// TIA Portal project "039_fw41" (V21)

(* hardware
DEVICE "PLC_1"  S7-1500 station
   slot 0: "Rail_0"  Rack  6ES7 590-1***0-0AA0
   slot 1: "PLC_1"  CPU 1516-3 PN/DP  6ES7 516-3AP03-0AB0  V4.1
      slot 3: "CPU display_1"  6ES7591-1BA00-0AA0
      slot 32768: "PROFINET interface_1"  X1
         slot 32769: "Port_1"  X1 P1
         slot 32770: "Port_2"  X1 P2
      slot 33024: "PROFINET interface_2"  X2
         slot 33025: "Port_1"  X2 P1
      slot 33280: "DP interface_1"  X3
      slot 34817: "Virtual CP interface port_1"  Virtual CP interface port  Virtual CP interface port FW V4.1
*)

// ===== PLC "PLC_1"  CPU 1516-3 PN/DP =====

DATA_BLOCK "DB_Arr"   // DB1
{ S7_Optimized_Access := 'FALSE' }
   VAR
      "a" : Array[0..9] of Int;
      "b" : Array[0..9] of Int;
      w : Array[0..3] of Word;
      r : Array[0..3] of Real;
      "by" : Array[0..7] of Byte;
      bits : Array[0..15] of Bool;
   END_VAR
BEGIN
END_DATA_BLOCK

FUNCTION_BLOCK "FX_Lad_103"   // FB1, LAD
{ S7_Optimized_Access := 'TRUE' }
VERSION : 0.1
   VAR_INPUT
      "a" : Bool;
      "b" : Bool;
      c : Bool;
      ia : Int;
      ib : Int;
      ic : Int;
      da : DInt;
      db : DInt;
      ra : Real;
      rb : Real;
      wa : Word;
      wb : Word;
      dwa : DWord;
      ba : Byte;
      ta : Time;
      tb : Time;
      s1 : String;
      s2 : String;
   END_VAR
   VAR_OUTPUT
      q : Bool;
      q2 : Bool;
      io : Int;
      io2 : Int;
      dout : DInt;
      rout : Real;
      wout : Word;
      dwout : DWord;
      bout : Byte;
      tout : Time;
      sout : String;
   END_VAR
   VAR_IN_OUT
      x_bool : Bool;
      x_uint : UInt;
      arr : Array[0..9] of Int;
      barr : Array[0..7] of Bool;
      iinout : Int;
   END_VAR
   VAR
      ton1 : TON_TIME;
      tof1 : TOF_TIME;
      tp1 : TP_TIME;
      tonr1 : TONR_TIME;
      ctu1 : CTU_INT;
      ctd1 : CTD_INT;
      ctud1 : CTUD_INT;
      rtrig1 : R_TRIG;
      ftrig1 : F_TRIG;
      edge1 : Bool;
      edge2 : Bool;
      stat1 : Bool;
      stat2 : Bool;
      stati : Int;
   END_VAR
   VAR_TEMP
      t1 : Bool;
      t2 : Bool;
      ti : Int;
      td : DInt;
      tr : Real;
      tw : Word;
      tt : Time;
      var1 : Variant;
   END_VAR
BEGIN

REGION Network 1: ---| |--- - Normally open contact
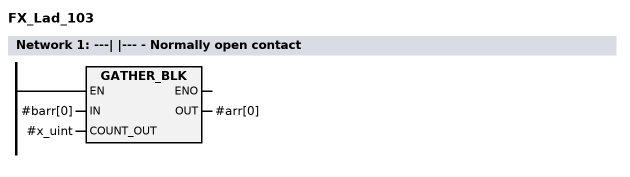
   GATHER_BLK(IN := #barr[0], COUNT_OUT := #x_uint, OUT => #arr[0]);
END_REGION
END_FUNCTION_BLOCK

FUNCTION_BLOCK "FX_TP2"   // FB2, LAD
{ S7_Optimized_Access := 'TRUE' }
VERSION : 0.1
   VAR_INPUT
      "a" : Bool;
      "b" : Bool;
      c : Bool;
      ia : Int;
      ib : Int;
      ic : Int;
      da : DInt;
      db : DInt;
      ra : Real;
      rb : Real;
      wa : Word;
      wb : Word;
      dwa : DWord;
      ba : Byte;
      ta : Time;
      tb : Time;
      s1 : String;
      s2 : String;
   END_VAR
   VAR_OUTPUT
      q : Bool;
      q2 : Bool;
      io : Int;
      io2 : Int;
      dout : DInt;
      rout : Real;
      wout : Word;
      dwout : DWord;
      bout : Byte;
      tout : Time;
      sout : String;
   END_VAR
   VAR_IN_OUT
      arr : Array[0..9] of Int;
      barr : Array[0..7] of Bool;
      iinout : Int;
   END_VAR
   VAR
      ton1 : TON_TIME;
      tof1 : TOF_TIME;
      tp1 : TP_TIME;
      tonr1 : TONR_TIME;
      ctu1 : CTU_INT;
      ctd1 : CTD_INT;
      ctud1 : CTUD_INT;
      rtrig1 : R_TRIG;
      ftrig1 : F_TRIG;
      edge1 : Bool;
      edge2 : Bool;
      stat1 : Bool;
      stat2 : Bool;
      stati : Int;
   END_VAR
   VAR_TEMP
      t1 : Bool;
      t2 : Bool;
      ti : Int;
      td : DInt;
      tr : Real;
      tw : Word;
      tt : Time;
      var1 : Variant;
   END_VAR
BEGIN

REGION Network 1: ---| |--- - Normally open contact
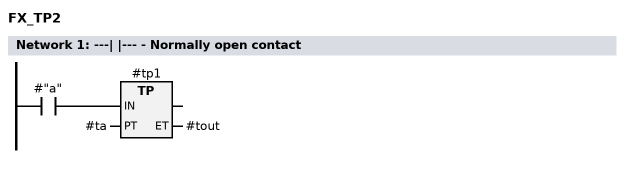
   #tp1(IN := #"a", PT := #ta, ET => #tout);   // TP
END_REGION
END_FUNCTION_BLOCK

FUNCTION_BLOCK "FX_Lad_024"   // FB3, LAD
{ S7_Optimized_Access := 'TRUE' }
VERSION : 0.1
   VAR_INPUT
      "a" : Bool;
      "b" : Bool;
      c : Bool;
      ia : Int;
      ib : Int;
      ic : Int;
      da : DInt;
      db : DInt;
      ra : Real;
      rb : Real;
      wa : Word;
      wb : Word;
      dwa : DWord;
      ba : Byte;
      ta : Time;
      tb : Time;
      s1 : String;
      s2 : String;
   END_VAR
   VAR_OUTPUT
      q : Bool;
      q2 : Bool;
      io : Int;
      io2 : Int;
      dout : DInt;
      rout : Real;
      wout : Word;
      dwout : DWord;
      bout : Byte;
      tout : Time;
      sout : String;
   END_VAR
   VAR_IN_OUT
      arr : Array[0..9] of Int;
      barr : Array[0..7] of Bool;
      iinout : Int;
   END_VAR
   VAR
      ton1 : TON_TIME;
      tof1 : TOF_TIME;
      tp1 : TP_TIME;
      tonr1 : TONR_TIME;
      ctu1 : CTU_INT;
      ctd1 : CTD_INT;
      ctud1 : CTUD_INT;
      rtrig1 : R_TRIG;
      ftrig1 : F_TRIG;
      edge1 : Bool;
      edge2 : Bool;
      stat1 : Bool;
      stat2 : Bool;
      stati : Int;
   END_VAR
   VAR_TEMP
      t1 : Bool;
      t2 : Bool;
      ti : Int;
      td : DInt;
      tr : Real;
      tw : Word;
      tt : Time;
      var1 : Variant;
   END_VAR
BEGIN

REGION Network 1: ---| |--- - Normally open contact
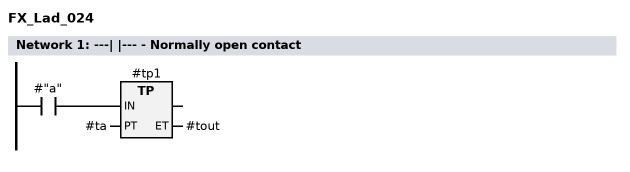
   #tp1(IN := #"a", PT := #ta, ET => #tout);   // TP
END_REGION
END_FUNCTION_BLOCK

FUNCTION_BLOCK "FX_Lad_025"   // FB4, LAD
{ S7_Optimized_Access := 'TRUE' }
VERSION : 0.1
   VAR_INPUT
      "a" : Bool;
      "b" : Bool;
      c : Bool;
      ia : Int;
      ib : Int;
      ic : Int;
      da : DInt;
      db : DInt;
      ra : Real;
      rb : Real;
      wa : Word;
      wb : Word;
      dwa : DWord;
      ba : Byte;
      ta : Time;
      tb : Time;
      s1 : String;
      s2 : String;
   END_VAR
   VAR_OUTPUT
      q : Bool;
      q2 : Bool;
      io : Int;
      io2 : Int;
      dout : DInt;
      rout : Real;
      wout : Word;
      dwout : DWord;
      bout : Byte;
      tout : Time;
      sout : String;
   END_VAR
   VAR_IN_OUT
      arr : Array[0..9] of Int;
      barr : Array[0..7] of Bool;
      iinout : Int;
   END_VAR
   VAR
      ton1 : TON_TIME;
      tof1 : TOF_TIME;
      tp1 : TP_TIME;
      tonr1 : TONR_TIME;
      ctu1 : CTU_INT;
      ctd1 : CTD_INT;
      ctud1 : CTUD_INT;
      rtrig1 : R_TRIG;
      ftrig1 : F_TRIG;
      edge1 : Bool;
      edge2 : Bool;
      stat1 : Bool;
      stat2 : Bool;
      stati : Int;
   END_VAR
   VAR_TEMP
      t1 : Bool;
      t2 : Bool;
      ti : Int;
      td : DInt;
      tr : Real;
      tw : Word;
      tt : Time;
      var1 : Variant;
   END_VAR
BEGIN

REGION Network 1: ---| |--- - Normally open contact
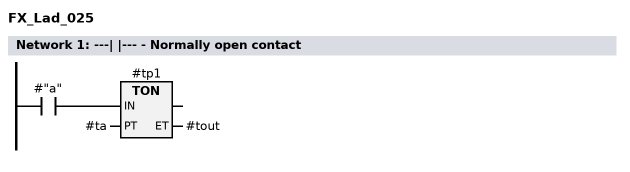
   #tp1(IN := #"a", PT := #ta, ET => #tout);   // TON
END_REGION
END_FUNCTION_BLOCK

FUNCTION_BLOCK "FX_Lad_026"   // FB5, LAD
{ S7_Optimized_Access := 'TRUE' }
VERSION : 0.1
   VAR_INPUT
      "a" : Bool;
      "b" : Bool;
      c : Bool;
      ia : Int;
      ib : Int;
      ic : Int;
      da : DInt;
      db : DInt;
      ra : Real;
      rb : Real;
      wa : Word;
      wb : Word;
      dwa : DWord;
      ba : Byte;
      ta : Time;
      tb : Time;
      s1 : String;
      s2 : String;
   END_VAR
   VAR_OUTPUT
      q : Bool;
      q2 : Bool;
      io : Int;
      io2 : Int;
      dout : DInt;
      rout : Real;
      wout : Word;
      dwout : DWord;
      bout : Byte;
      tout : Time;
      sout : String;
   END_VAR
   VAR_IN_OUT
      arr : Array[0..9] of Int;
      barr : Array[0..7] of Bool;
      iinout : Int;
   END_VAR
   VAR
      ton1 : TON_TIME;
      tof1 : TOF_TIME;
      tp1 : TP_TIME;
      tonr1 : TONR_TIME;
      ctu1 : CTU_INT;
      ctd1 : CTD_INT;
      ctud1 : CTUD_INT;
      rtrig1 : R_TRIG;
      ftrig1 : F_TRIG;
      edge1 : Bool;
      edge2 : Bool;
      stat1 : Bool;
      stat2 : Bool;
      stati : Int;
   END_VAR
   VAR_TEMP
      t1 : Bool;
      t2 : Bool;
      ti : Int;
      td : DInt;
      tr : Real;
      tw : Word;
      tt : Time;
      var1 : Variant;
   END_VAR
BEGIN

REGION Network 1: ---| |--- - Normally open contact
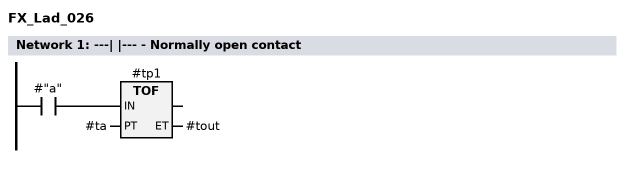
   #tp1(IN := #"a", PT := #ta, ET => #tout);   // TOF
END_REGION
END_FUNCTION_BLOCK

FUNCTION_BLOCK "FX_Lad_027"   // FB6, LAD
{ S7_Optimized_Access := 'TRUE' }
VERSION : 0.1
   VAR_INPUT
      "a" : Bool;
      "b" : Bool;
      c : Bool;
      ia : Int;
      ib : Int;
      ic : Int;
      da : DInt;
      db : DInt;
      ra : Real;
      rb : Real;
      wa : Word;
      wb : Word;
      dwa : DWord;
      ba : Byte;
      ta : Time;
      tb : Time;
      s1 : String;
      s2 : String;
   END_VAR
   VAR_OUTPUT
      q : Bool;
      q2 : Bool;
      io : Int;
      io2 : Int;
      dout : DInt;
      rout : Real;
      wout : Word;
      dwout : DWord;
      bout : Byte;
      tout : Time;
      sout : String;
   END_VAR
   VAR_IN_OUT
      arr : Array[0..9] of Int;
      barr : Array[0..7] of Bool;
      iinout : Int;
   END_VAR
   VAR
      ton1 : TON_TIME;
      tof1 : TOF_TIME;
      tp1 : TP_TIME;
      tonr1 : TONR_TIME;
      ctu1 : CTU_INT;
      ctd1 : CTD_INT;
      ctud1 : CTUD_INT;
      rtrig1 : R_TRIG;
      ftrig1 : F_TRIG;
      edge1 : Bool;
      edge2 : Bool;
      stat1 : Bool;
      stat2 : Bool;
      stati : Int;
   END_VAR
   VAR_TEMP
      t1 : Bool;
      t2 : Bool;
      ti : Int;
      td : DInt;
      tr : Real;
      tw : Word;
      tt : Time;
      var1 : Variant;
   END_VAR
BEGIN

REGION Network 1: ---| |--- - Normally open contact
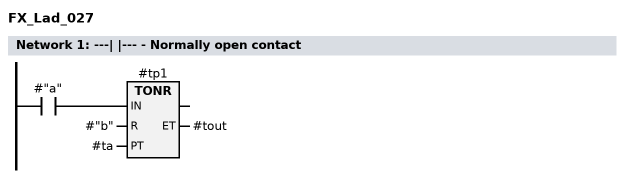
   #tp1(IN := #"a", R := #"b", PT := #ta, ET => #tout);   // TONR
END_REGION
END_FUNCTION_BLOCK

FUNCTION_BLOCK "FX_Lad_ex003"   // FB7, LAD
{ S7_Optimized_Access := 'TRUE' }
VERSION : 0.1
   VAR_INPUT
      "a" : Bool;
      "b" : Bool;
      c : Bool;
      ia : Int;
      ib : Int;
      ic : Int;
      da : DInt;
      db : DInt;
      ra : Real;
      rb : Real;
      wa : Word;
      wb : Word;
      dwa : DWord;
      ba : Byte;
      ta : Time;
      tb : Time;
      s1 : String;
      s2 : String;
   END_VAR
   VAR_OUTPUT
      q : Bool;
      q2 : Bool;
      io : Int;
      io2 : Int;
      dout : DInt;
      rout : Real;
      wout : Word;
      dwout : DWord;
      bout : Byte;
      tout : Time;
      sout : String;
   END_VAR
   VAR_IN_OUT
      x_time : Time;
      arr : Array[0..9] of Int;
      barr : Array[0..7] of Bool;
      iinout : Int;
   END_VAR
   VAR
      ton1 : TON_TIME;
      tof1 : TOF_TIME;
      tp1 : TP_TIME;
      tonr1 : TONR_TIME;
      ctu1 : CTU_INT;
      ctd1 : CTD_INT;
      ctud1 : CTUD_INT;
      rtrig1 : R_TRIG;
      ftrig1 : F_TRIG;
      edge1 : Bool;
      edge2 : Bool;
      stat1 : Bool;
      stat2 : Bool;
      stati : Int;
   END_VAR
   VAR_TEMP
      t1 : Bool;
      t2 : Bool;
      ti : Int;
      td : DInt;
      tr : Real;
      tw : Word;
      tt : Time;
      var1 : Variant;
   END_VAR
BEGIN

REGION Network 1: ---| |--- - Normally open contact
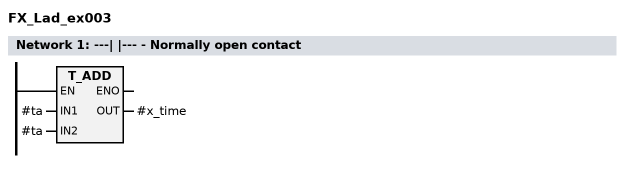
   #x_time := T_ADD(IN1 := #ta, IN2 := #ta);
END_REGION
END_FUNCTION_BLOCK

FUNCTION_BLOCK "FX_Lad_ex004"   // FB8, LAD
{ S7_Optimized_Access := 'TRUE' }
VERSION : 0.1
   VAR_INPUT
      "a" : Bool;
      "b" : Bool;
      c : Bool;
      ia : Int;
      ib : Int;
      ic : Int;
      da : DInt;
      db : DInt;
      ra : Real;
      rb : Real;
      wa : Word;
      wb : Word;
      dwa : DWord;
      ba : Byte;
      ta : Time;
      tb : Time;
      s1 : String;
      s2 : String;
   END_VAR
   VAR_OUTPUT
      q : Bool;
      q2 : Bool;
      io : Int;
      io2 : Int;
      dout : DInt;
      rout : Real;
      wout : Word;
      dwout : DWord;
      bout : Byte;
      tout : Time;
      sout : String;
   END_VAR
   VAR_IN_OUT
      x_time : Time;
      arr : Array[0..9] of Int;
      barr : Array[0..7] of Bool;
      iinout : Int;
   END_VAR
   VAR
      ton1 : TON_TIME;
      tof1 : TOF_TIME;
      tp1 : TP_TIME;
      tonr1 : TONR_TIME;
      ctu1 : CTU_INT;
      ctd1 : CTD_INT;
      ctud1 : CTUD_INT;
      rtrig1 : R_TRIG;
      ftrig1 : F_TRIG;
      edge1 : Bool;
      edge2 : Bool;
      stat1 : Bool;
      stat2 : Bool;
      stati : Int;
   END_VAR
   VAR_TEMP
      t1 : Bool;
      t2 : Bool;
      ti : Int;
      td : DInt;
      tr : Real;
      tw : Word;
      tt : Time;
      var1 : Variant;
   END_VAR
BEGIN

REGION Network 1: ---| |--- - Normally open contact
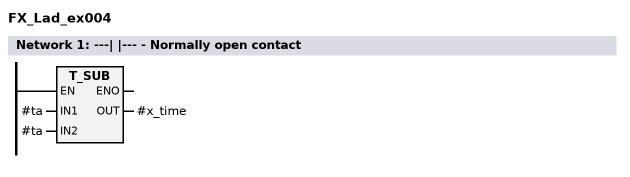
   #x_time := T_SUB(IN1 := #ta, IN2 := #ta);
END_REGION
END_FUNCTION_BLOCK

FUNCTION_BLOCK "FX_Lad_ex018"   // FB9, LAD
{ S7_Optimized_Access := 'TRUE' }
VERSION : 0.1
   VAR_INPUT
      "a" : Bool;
      "b" : Bool;
      c : Bool;
      ia : Int;
      ib : Int;
      ic : Int;
      da : DInt;
      db : DInt;
      ra : Real;
      rb : Real;
      wa : Word;
      wb : Word;
      dwa : DWord;
      ba : Byte;
      ta : Time;
      tb : Time;
      s1 : String;
      s2 : String;
   END_VAR
   VAR_OUTPUT
      q : Bool;
      q2 : Bool;
      io : Int;
      io2 : Int;
      dout : DInt;
      rout : Real;
      wout : Word;
      dwout : DWord;
      bout : Byte;
      tout : Time;
      sout : String;
   END_VAR
   VAR_IN_OUT
      arr : Array[0..9] of Int;
      barr : Array[0..7] of Bool;
      iinout : Int;
   END_VAR
   VAR
      ton1 : TON_TIME;
      tof1 : TOF_TIME;
      tp1 : TP_TIME;
      tonr1 : TONR_TIME;
      ctu1 : CTU_INT;
      ctd1 : CTD_INT;
      ctud1 : CTUD_INT;
      rtrig1 : R_TRIG;
      ftrig1 : F_TRIG;
      edge1 : Bool;
      edge2 : Bool;
      stat1 : Bool;
      stat2 : Bool;
      stati : Int;
   END_VAR
   VAR_TEMP
      t1 : Bool;
      t2 : Bool;
      ti : Int;
      td : DInt;
      tr : Real;
      tw : Word;
      tt : Time;
      var1 : Variant;
   END_VAR
BEGIN

REGION Network 1: ---| |--- - Normally open contact
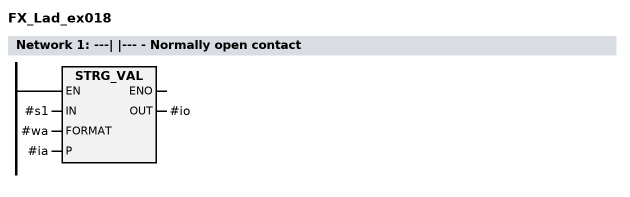
   STRG_VAL(IN := #s1, FORMAT := #wa, P := #ia, OUT => #io);
END_REGION
END_FUNCTION_BLOCK

FUNCTION_BLOCK "FX_Lad_ex019"   // FB10, LAD
{ S7_Optimized_Access := 'TRUE' }
VERSION : 0.1
   VAR_INPUT
      "a" : Bool;
      "b" : Bool;
      c : Bool;
      ia : Int;
      ib : Int;
      ic : Int;
      da : DInt;
      db : DInt;
      ra : Real;
      rb : Real;
      wa : Word;
      wb : Word;
      dwa : DWord;
      ba : Byte;
      ta : Time;
      tb : Time;
      s1 : String;
      s2 : String;
   END_VAR
   VAR_OUTPUT
      q : Bool;
      q2 : Bool;
      io : Int;
      io2 : Int;
      dout : DInt;
      rout : Real;
      wout : Word;
      dwout : DWord;
      bout : Byte;
      tout : Time;
      sout : String;
   END_VAR
   VAR_IN_OUT
      arr : Array[0..9] of Int;
      barr : Array[0..7] of Bool;
      iinout : Int;
   END_VAR
   VAR
      ton1 : TON_TIME;
      tof1 : TOF_TIME;
      tp1 : TP_TIME;
      tonr1 : TONR_TIME;
      ctu1 : CTU_INT;
      ctd1 : CTD_INT;
      ctud1 : CTUD_INT;
      rtrig1 : R_TRIG;
      ftrig1 : F_TRIG;
      edge1 : Bool;
      edge2 : Bool;
      stat1 : Bool;
      stat2 : Bool;
      stati : Int;
   END_VAR
   VAR_TEMP
      t1 : Bool;
      t2 : Bool;
      ti : Int;
      td : DInt;
      tr : Real;
      tw : Word;
      tt : Time;
      var1 : Variant;
   END_VAR
BEGIN

REGION Network 1: ---| |--- - Normally open contact
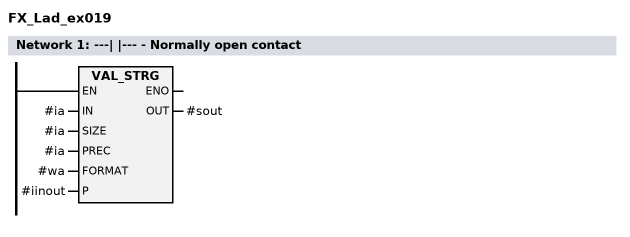
   VAL_STRG(IN := #ia, SIZE := #ia, PREC := #ia, FORMAT := #wa, P := #iinout, OUT => #sout);
END_REGION
END_FUNCTION_BLOCK

FUNCTION_BLOCK "FX_Lad_ex021"   // FB11, LAD
{ S7_Optimized_Access := 'TRUE' }
VERSION : 0.1
   VAR_INPUT
      "a" : Bool;
      "b" : Bool;
      c : Bool;
      ia : Int;
      ib : Int;
      ic : Int;
      da : DInt;
      db : DInt;
      ra : Real;
      rb : Real;
      wa : Word;
      wb : Word;
      dwa : DWord;
      ba : Byte;
      ta : Time;
      tb : Time;
      s1 : String;
      s2 : String;
   END_VAR
   VAR_OUTPUT
      q : Bool;
      q2 : Bool;
      io : Int;
      io2 : Int;
      dout : DInt;
      rout : Real;
      wout : Word;
      dwout : DWord;
      bout : Byte;
      tout : Time;
      sout : String;
   END_VAR
   VAR_IN_OUT
      x_variant : Variant;
      arr : Array[0..9] of Int;
      barr : Array[0..7] of Bool;
      iinout : Int;
   END_VAR
   VAR
      ton1 : TON_TIME;
      tof1 : TOF_TIME;
      tp1 : TP_TIME;
      tonr1 : TONR_TIME;
      ctu1 : CTU_INT;
      ctd1 : CTD_INT;
      ctud1 : CTUD_INT;
      rtrig1 : R_TRIG;
      ftrig1 : F_TRIG;
      edge1 : Bool;
      edge2 : Bool;
      stat1 : Bool;
      stat2 : Bool;
      stati : Int;
   END_VAR
   VAR_TEMP
      t1 : Bool;
      t2 : Bool;
      ti : Int;
      td : DInt;
      tr : Real;
      tw : Word;
      tt : Time;
      var1 : Variant;
   END_VAR
BEGIN

REGION Network 1: ---| |--- - Normally open contact
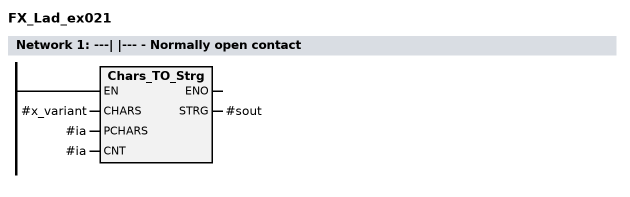
   // no SCL statement known for Chars_TO_Strg: written as a call
   Chars_TO_Strg(Chars := #x_variant, pChars := #ia, Cnt := #ia, Strg => #sout);
END_REGION
END_FUNCTION_BLOCK

FUNCTION_BLOCK "FX_Lad_ex027"   // FB12, LAD
{ S7_Optimized_Access := 'TRUE' }
VERSION : 0.1
   VAR_INPUT
      "a" : Bool;
      "b" : Bool;
      c : Bool;
      ia : Int;
      ib : Int;
      ic : Int;
      da : DInt;
      db : DInt;
      ra : Real;
      rb : Real;
      wa : Word;
      wb : Word;
      dwa : DWord;
      ba : Byte;
      ta : Time;
      tb : Time;
      s1 : String;
      s2 : String;
   END_VAR
   VAR_OUTPUT
      q : Bool;
      q2 : Bool;
      io : Int;
      io2 : Int;
      dout : DInt;
      rout : Real;
      wout : Word;
      dwout : DWord;
      bout : Byte;
      tout : Time;
      sout : String;
   END_VAR
   VAR_IN_OUT
      arr : Array[0..9] of Int;
      barr : Array[0..7] of Bool;
      iinout : Int;
   END_VAR
   VAR
      ton1 : TON_TIME;
      tof1 : TOF_TIME;
      tp1 : TP_TIME;
      tonr1 : TONR_TIME;
      ctu1 : CTU_INT;
      ctd1 : CTD_INT;
      ctud1 : CTUD_INT;
      rtrig1 : R_TRIG;
      ftrig1 : F_TRIG;
      edge1 : Bool;
      edge2 : Bool;
      stat1 : Bool;
      stat2 : Bool;
      stati : Int;
   END_VAR
   VAR_TEMP
      t1 : Bool;
      t2 : Bool;
      ti : Int;
      td : DInt;
      tr : Real;
      tw : Word;
      tt : Time;
      var1 : Variant;
   END_VAR
BEGIN

REGION Network 1: ---| |--- - Normally open contact
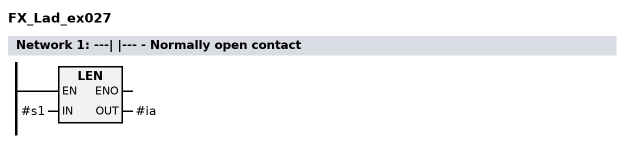
   #ia := LEN(IN := #s1);
END_REGION
END_FUNCTION_BLOCK

FUNCTION_BLOCK "FX_Lad_ex028"   // FB13, LAD
{ S7_Optimized_Access := 'TRUE' }
VERSION : 0.1
   VAR_INPUT
      "a" : Bool;
      "b" : Bool;
      c : Bool;
      ia : Int;
      ib : Int;
      ic : Int;
      da : DInt;
      db : DInt;
      ra : Real;
      rb : Real;
      wa : Word;
      wb : Word;
      dwa : DWord;
      ba : Byte;
      ta : Time;
      tb : Time;
      s1 : String;
      s2 : String;
   END_VAR
   VAR_OUTPUT
      q : Bool;
      q2 : Bool;
      io : Int;
      io2 : Int;
      dout : DInt;
      rout : Real;
      wout : Word;
      dwout : DWord;
      bout : Byte;
      tout : Time;
      sout : String;
   END_VAR
   VAR_IN_OUT
      arr : Array[0..9] of Int;
      barr : Array[0..7] of Bool;
      iinout : Int;
   END_VAR
   VAR
      ton1 : TON_TIME;
      tof1 : TOF_TIME;
      tp1 : TP_TIME;
      tonr1 : TONR_TIME;
      ctu1 : CTU_INT;
      ctd1 : CTD_INT;
      ctud1 : CTUD_INT;
      rtrig1 : R_TRIG;
      ftrig1 : F_TRIG;
      edge1 : Bool;
      edge2 : Bool;
      stat1 : Bool;
      stat2 : Bool;
      stati : Int;
   END_VAR
   VAR_TEMP
      t1 : Bool;
      t2 : Bool;
      ti : Int;
      td : DInt;
      tr : Real;
      tw : Word;
      tt : Time;
      var1 : Variant;
   END_VAR
BEGIN

REGION Network 1: ---| |--- - Normally open contact
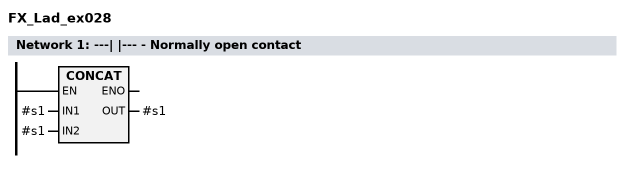
   #s1 := CONCAT(IN1 := #s1, IN2 := #s1);
END_REGION
END_FUNCTION_BLOCK

FUNCTION_BLOCK "FX_Lad_ex029"   // FB14, LAD
{ S7_Optimized_Access := 'TRUE' }
VERSION : 0.1
   VAR_INPUT
      "a" : Bool;
      "b" : Bool;
      c : Bool;
      ia : Int;
      ib : Int;
      ic : Int;
      da : DInt;
      db : DInt;
      ra : Real;
      rb : Real;
      wa : Word;
      wb : Word;
      dwa : DWord;
      ba : Byte;
      ta : Time;
      tb : Time;
      s1 : String;
      s2 : String;
   END_VAR
   VAR_OUTPUT
      q : Bool;
      q2 : Bool;
      io : Int;
      io2 : Int;
      dout : DInt;
      rout : Real;
      wout : Word;
      dwout : DWord;
      bout : Byte;
      tout : Time;
      sout : String;
   END_VAR
   VAR_IN_OUT
      arr : Array[0..9] of Int;
      barr : Array[0..7] of Bool;
      iinout : Int;
   END_VAR
   VAR
      ton1 : TON_TIME;
      tof1 : TOF_TIME;
      tp1 : TP_TIME;
      tonr1 : TONR_TIME;
      ctu1 : CTU_INT;
      ctd1 : CTD_INT;
      ctud1 : CTUD_INT;
      rtrig1 : R_TRIG;
      ftrig1 : F_TRIG;
      edge1 : Bool;
      edge2 : Bool;
      stat1 : Bool;
      stat2 : Bool;
      stati : Int;
   END_VAR
   VAR_TEMP
      t1 : Bool;
      t2 : Bool;
      ti : Int;
      td : DInt;
      tr : Real;
      tw : Word;
      tt : Time;
      var1 : Variant;
   END_VAR
BEGIN

REGION Network 1: ---| |--- - Normally open contact
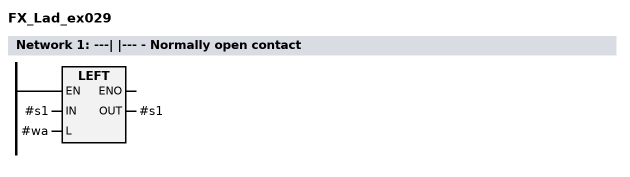
   #s1 := LEFT(IN := #s1, L := #wa);
END_REGION
END_FUNCTION_BLOCK

FUNCTION_BLOCK "FX_Lad_ex030"   // FB15, LAD
{ S7_Optimized_Access := 'TRUE' }
VERSION : 0.1
   VAR_INPUT
      "a" : Bool;
      "b" : Bool;
      c : Bool;
      ia : Int;
      ib : Int;
      ic : Int;
      da : DInt;
      db : DInt;
      ra : Real;
      rb : Real;
      wa : Word;
      wb : Word;
      dwa : DWord;
      ba : Byte;
      ta : Time;
      tb : Time;
      s1 : String;
      s2 : String;
   END_VAR
   VAR_OUTPUT
      q : Bool;
      q2 : Bool;
      io : Int;
      io2 : Int;
      dout : DInt;
      rout : Real;
      wout : Word;
      dwout : DWord;
      bout : Byte;
      tout : Time;
      sout : String;
   END_VAR
   VAR_IN_OUT
      arr : Array[0..9] of Int;
      barr : Array[0..7] of Bool;
      iinout : Int;
   END_VAR
   VAR
      ton1 : TON_TIME;
      tof1 : TOF_TIME;
      tp1 : TP_TIME;
      tonr1 : TONR_TIME;
      ctu1 : CTU_INT;
      ctd1 : CTD_INT;
      ctud1 : CTUD_INT;
      rtrig1 : R_TRIG;
      ftrig1 : F_TRIG;
      edge1 : Bool;
      edge2 : Bool;
      stat1 : Bool;
      stat2 : Bool;
      stati : Int;
   END_VAR
   VAR_TEMP
      t1 : Bool;
      t2 : Bool;
      ti : Int;
      td : DInt;
      tr : Real;
      tw : Word;
      tt : Time;
      var1 : Variant;
   END_VAR
BEGIN

REGION Network 1: ---| |--- - Normally open contact
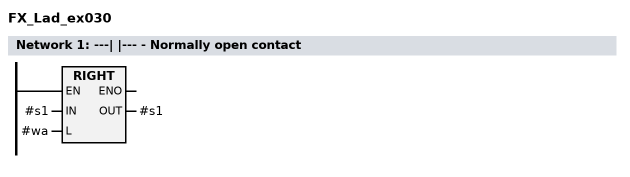
   #s1 := RIGHT(IN := #s1, L := #wa);
END_REGION
END_FUNCTION_BLOCK

FUNCTION_BLOCK "FX_Lad_ex031"   // FB16, LAD
{ S7_Optimized_Access := 'TRUE' }
VERSION : 0.1
   VAR_INPUT
      "a" : Bool;
      "b" : Bool;
      c : Bool;
      ia : Int;
      ib : Int;
      ic : Int;
      da : DInt;
      db : DInt;
      ra : Real;
      rb : Real;
      wa : Word;
      wb : Word;
      dwa : DWord;
      ba : Byte;
      ta : Time;
      tb : Time;
      s1 : String;
      s2 : String;
   END_VAR
   VAR_OUTPUT
      q : Bool;
      q2 : Bool;
      io : Int;
      io2 : Int;
      dout : DInt;
      rout : Real;
      wout : Word;
      dwout : DWord;
      bout : Byte;
      tout : Time;
      sout : String;
   END_VAR
   VAR_IN_OUT
      arr : Array[0..9] of Int;
      barr : Array[0..7] of Bool;
      iinout : Int;
   END_VAR
   VAR
      ton1 : TON_TIME;
      tof1 : TOF_TIME;
      tp1 : TP_TIME;
      tonr1 : TONR_TIME;
      ctu1 : CTU_INT;
      ctd1 : CTD_INT;
      ctud1 : CTUD_INT;
      rtrig1 : R_TRIG;
      ftrig1 : F_TRIG;
      edge1 : Bool;
      edge2 : Bool;
      stat1 : Bool;
      stat2 : Bool;
      stati : Int;
   END_VAR
   VAR_TEMP
      t1 : Bool;
      t2 : Bool;
      ti : Int;
      td : DInt;
      tr : Real;
      tw : Word;
      tt : Time;
      var1 : Variant;
   END_VAR
BEGIN

REGION Network 1: ---| |--- - Normally open contact
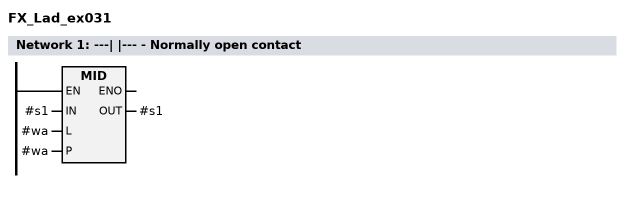
   #s1 := MID(IN := #s1, L := #wa, P := #wa);
END_REGION
END_FUNCTION_BLOCK

FUNCTION_BLOCK "FX_Lad_ex032"   // FB17, LAD
{ S7_Optimized_Access := 'TRUE' }
VERSION : 0.1
   VAR_INPUT
      "a" : Bool;
      "b" : Bool;
      c : Bool;
      ia : Int;
      ib : Int;
      ic : Int;
      da : DInt;
      db : DInt;
      ra : Real;
      rb : Real;
      wa : Word;
      wb : Word;
      dwa : DWord;
      ba : Byte;
      ta : Time;
      tb : Time;
      s1 : String;
      s2 : String;
   END_VAR
   VAR_OUTPUT
      q : Bool;
      q2 : Bool;
      io : Int;
      io2 : Int;
      dout : DInt;
      rout : Real;
      wout : Word;
      dwout : DWord;
      bout : Byte;
      tout : Time;
      sout : String;
   END_VAR
   VAR_IN_OUT
      arr : Array[0..9] of Int;
      barr : Array[0..7] of Bool;
      iinout : Int;
   END_VAR
   VAR
      ton1 : TON_TIME;
      tof1 : TOF_TIME;
      tp1 : TP_TIME;
      tonr1 : TONR_TIME;
      ctu1 : CTU_INT;
      ctd1 : CTD_INT;
      ctud1 : CTUD_INT;
      rtrig1 : R_TRIG;
      ftrig1 : F_TRIG;
      edge1 : Bool;
      edge2 : Bool;
      stat1 : Bool;
      stat2 : Bool;
      stati : Int;
   END_VAR
   VAR_TEMP
      t1 : Bool;
      t2 : Bool;
      ti : Int;
      td : DInt;
      tr : Real;
      tw : Word;
      tt : Time;
      var1 : Variant;
   END_VAR
BEGIN

REGION Network 1: ---| |--- - Normally open contact
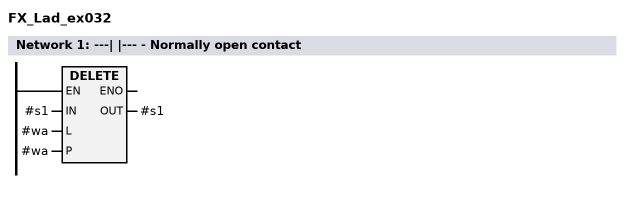
   #s1 := DELETE(IN := #s1, L := #wa, P := #wa);
END_REGION
END_FUNCTION_BLOCK

FUNCTION_BLOCK "FX_Lad_ex033"   // FB18, LAD
{ S7_Optimized_Access := 'TRUE' }
VERSION : 0.1
   VAR_INPUT
      "a" : Bool;
      "b" : Bool;
      c : Bool;
      ia : Int;
      ib : Int;
      ic : Int;
      da : DInt;
      db : DInt;
      ra : Real;
      rb : Real;
      wa : Word;
      wb : Word;
      dwa : DWord;
      ba : Byte;
      ta : Time;
      tb : Time;
      s1 : String;
      s2 : String;
   END_VAR
   VAR_OUTPUT
      q : Bool;
      q2 : Bool;
      io : Int;
      io2 : Int;
      dout : DInt;
      rout : Real;
      wout : Word;
      dwout : DWord;
      bout : Byte;
      tout : Time;
      sout : String;
   END_VAR
   VAR_IN_OUT
      arr : Array[0..9] of Int;
      barr : Array[0..7] of Bool;
      iinout : Int;
   END_VAR
   VAR
      ton1 : TON_TIME;
      tof1 : TOF_TIME;
      tp1 : TP_TIME;
      tonr1 : TONR_TIME;
      ctu1 : CTU_INT;
      ctd1 : CTD_INT;
      ctud1 : CTUD_INT;
      rtrig1 : R_TRIG;
      ftrig1 : F_TRIG;
      edge1 : Bool;
      edge2 : Bool;
      stat1 : Bool;
      stat2 : Bool;
      stati : Int;
   END_VAR
   VAR_TEMP
      t1 : Bool;
      t2 : Bool;
      ti : Int;
      td : DInt;
      tr : Real;
      tw : Word;
      tt : Time;
      var1 : Variant;
   END_VAR
BEGIN

REGION Network 1: ---| |--- - Normally open contact
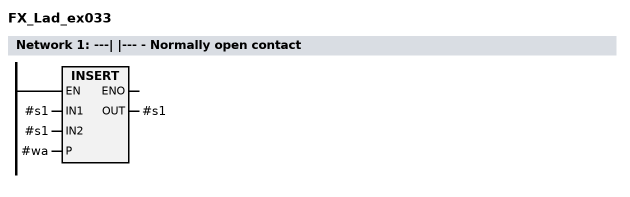
   #s1 := INSERT(IN1 := #s1, IN2 := #s1, P := #wa);
END_REGION
END_FUNCTION_BLOCK

FUNCTION_BLOCK "FX_Lad_ex034"   // FB19, LAD
{ S7_Optimized_Access := 'TRUE' }
VERSION : 0.1
   VAR_INPUT
      "a" : Bool;
      "b" : Bool;
      c : Bool;
      ia : Int;
      ib : Int;
      ic : Int;
      da : DInt;
      db : DInt;
      ra : Real;
      rb : Real;
      wa : Word;
      wb : Word;
      dwa : DWord;
      ba : Byte;
      ta : Time;
      tb : Time;
      s1 : String;
      s2 : String;
   END_VAR
   VAR_OUTPUT
      q : Bool;
      q2 : Bool;
      io : Int;
      io2 : Int;
      dout : DInt;
      rout : Real;
      wout : Word;
      dwout : DWord;
      bout : Byte;
      tout : Time;
      sout : String;
   END_VAR
   VAR_IN_OUT
      arr : Array[0..9] of Int;
      barr : Array[0..7] of Bool;
      iinout : Int;
   END_VAR
   VAR
      ton1 : TON_TIME;
      tof1 : TOF_TIME;
      tp1 : TP_TIME;
      tonr1 : TONR_TIME;
      ctu1 : CTU_INT;
      ctd1 : CTD_INT;
      ctud1 : CTUD_INT;
      rtrig1 : R_TRIG;
      ftrig1 : F_TRIG;
      edge1 : Bool;
      edge2 : Bool;
      stat1 : Bool;
      stat2 : Bool;
      stati : Int;
   END_VAR
   VAR_TEMP
      t1 : Bool;
      t2 : Bool;
      ti : Int;
      td : DInt;
      tr : Real;
      tw : Word;
      tt : Time;
      var1 : Variant;
   END_VAR
BEGIN

REGION Network 1: ---| |--- - Normally open contact
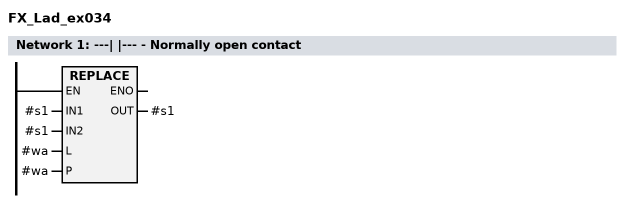
   #s1 := REPLACE(IN1 := #s1, IN2 := #s1, L := #wa, P := #wa);
END_REGION
END_FUNCTION_BLOCK

FUNCTION_BLOCK "FX_Lad_ex035"   // FB20, LAD
{ S7_Optimized_Access := 'TRUE' }
VERSION : 0.1
   VAR_INPUT
      "a" : Bool;
      "b" : Bool;
      c : Bool;
      ia : Int;
      ib : Int;
      ic : Int;
      da : DInt;
      db : DInt;
      ra : Real;
      rb : Real;
      wa : Word;
      wb : Word;
      dwa : DWord;
      ba : Byte;
      ta : Time;
      tb : Time;
      s1 : String;
      s2 : String;
   END_VAR
   VAR_OUTPUT
      q : Bool;
      q2 : Bool;
      io : Int;
      io2 : Int;
      dout : DInt;
      rout : Real;
      wout : Word;
      dwout : DWord;
      bout : Byte;
      tout : Time;
      sout : String;
   END_VAR
   VAR_IN_OUT
      arr : Array[0..9] of Int;
      barr : Array[0..7] of Bool;
      iinout : Int;
   END_VAR
   VAR
      ton1 : TON_TIME;
      tof1 : TOF_TIME;
      tp1 : TP_TIME;
      tonr1 : TONR_TIME;
      ctu1 : CTU_INT;
      ctd1 : CTD_INT;
      ctud1 : CTUD_INT;
      rtrig1 : R_TRIG;
      ftrig1 : F_TRIG;
      edge1 : Bool;
      edge2 : Bool;
      stat1 : Bool;
      stat2 : Bool;
      stati : Int;
   END_VAR
   VAR_TEMP
      t1 : Bool;
      t2 : Bool;
      ti : Int;
      td : DInt;
      tr : Real;
      tw : Word;
      tt : Time;
      var1 : Variant;
   END_VAR
BEGIN

REGION Network 1: ---| |--- - Normally open contact
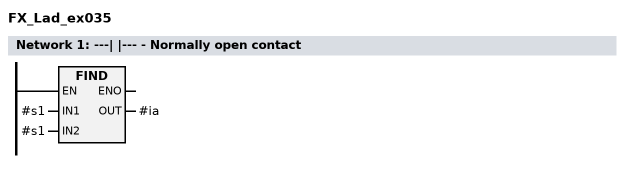
   #ia := FIND(IN1 := #s1, IN2 := #s1);
END_REGION
END_FUNCTION_BLOCK

FUNCTION_BLOCK "FX_Lad_ex159"   // FB21, LAD
{ S7_Optimized_Access := 'TRUE' }
VERSION : 0.1
   VAR_INPUT
      "a" : Bool;
      "b" : Bool;
      c : Bool;
      ia : Int;
      ib : Int;
      ic : Int;
      da : DInt;
      db : DInt;
      ra : Real;
      rb : Real;
      wa : Word;
      wb : Word;
      dwa : DWord;
      ba : Byte;
      ta : Time;
      tb : Time;
      s1 : String;
      s2 : String;
   END_VAR
   VAR_OUTPUT
      q : Bool;
      q2 : Bool;
      io : Int;
      io2 : Int;
      dout : DInt;
      rout : Real;
      wout : Word;
      dwout : DWord;
      bout : Byte;
      tout : Time;
      sout : String;
   END_VAR
   VAR_IN_OUT
      x_hw_any : Hw_Any;
      arr : Array[0..9] of Int;
      barr : Array[0..7] of Bool;
      iinout : Int;
   END_VAR
   VAR
      ton1 : TON_TIME;
      tof1 : TOF_TIME;
      tp1 : TP_TIME;
      tonr1 : TONR_TIME;
      ctu1 : CTU_INT;
      ctd1 : CTD_INT;
      ctud1 : CTUD_INT;
      rtrig1 : R_TRIG;
      ftrig1 : F_TRIG;
      edge1 : Bool;
      edge2 : Bool;
      stat1 : Bool;
      stat2 : Bool;
      stati : Int;
   END_VAR
   VAR_TEMP
      t1 : Bool;
      t2 : Bool;
      ti : Int;
      td : DInt;
      tr : Real;
      tw : Word;
      tt : Time;
      var1 : Variant;
   END_VAR
BEGIN

REGION Network 1: ---| |--- - Normally open contact
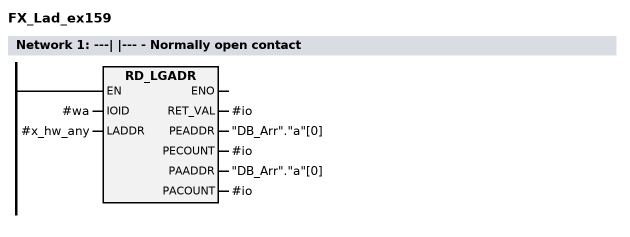
   // no checked SCL form for this network; see the picture
END_REGION
END_FUNCTION_BLOCK

FUNCTION_BLOCK "FB_Scl_sl001"   // FB22, SCL
{ S7_Optimized_Access := 'TRUE' }
VERSION : 0.1
   VAR_INPUT
      v_clk : Bool;
   END_VAR
   VAR_OUTPUT
      v_q : Bool;
   END_VAR
   VAR
      inst : R_TRIG;
   END_VAR
BEGIN
   #inst(CLK := #v_clk, Q => #v_q);
END_FUNCTION_BLOCK

FUNCTION_BLOCK "FB_Scl_sl003"   // FB23, SCL
{ S7_Optimized_Access := 'TRUE' }
VERSION : 0.1
   VAR_INPUT
      v_in : Bool;
      v_pt : Time;
   END_VAR
   VAR_OUTPUT
      v_q : Bool;
      v_et : Time;
   END_VAR
   VAR
      inst : TP_TIME;
   END_VAR
BEGIN
   #inst(IN := #v_in, PT := #v_pt, Q => #v_q, ET => #v_et);
END_FUNCTION_BLOCK

FUNCTION_BLOCK "FB_Scl_sl014"   // FB24, SCL
{ S7_Optimized_Access := 'TRUE' }
VERSION : 0.1
   VAR_INPUT
      v_cu : Bool;
      v_r : Bool;
      v_pv : Int;
   END_VAR
   VAR_OUTPUT
      v_q : Bool;
      v_cv : Char;
   END_VAR
   VAR
      inst : CTU_INT;
   END_VAR
BEGIN
   #inst(CU := #v_cu, R := #v_r, PV := #v_pv, Q => #v_q, CV => #v_cv);
END_FUNCTION_BLOCK

FUNCTION_BLOCK "FB_Scl_sl002"   // FB25, SCL
{ S7_Optimized_Access := 'TRUE' }
VERSION : 0.1
   VAR_INPUT
      v_clk : Bool;
   END_VAR
   VAR_OUTPUT
      v_q : Bool;
   END_VAR
   VAR
      inst : F_TRIG;
   END_VAR
BEGIN
   #inst(CLK := #v_clk, Q => #v_q);
END_FUNCTION_BLOCK

FUNCTION_BLOCK "FB_Scl_sl004"   // FB26, SCL
{ S7_Optimized_Access := 'TRUE' }
VERSION : 0.1
   VAR_INPUT
      v_in : Bool;
      v_pt : Time;
   END_VAR
   VAR_OUTPUT
      v_q : Bool;
      v_et : Time;
   END_VAR
   VAR
      inst : TON_TIME;
   END_VAR
BEGIN
   #inst(IN := #v_in, PT := #v_pt, Q => #v_q, ET => #v_et);
END_FUNCTION_BLOCK

FUNCTION_BLOCK "FB_Scl_sl005"   // FB27, SCL
{ S7_Optimized_Access := 'TRUE' }
VERSION : 0.1
   VAR_INPUT
      v_in : Bool;
      v_pt : Time;
   END_VAR
   VAR_OUTPUT
      v_q : Bool;
      v_et : Time;
   END_VAR
   VAR
      inst : TOF_TIME;
   END_VAR
BEGIN
   #inst(IN := #v_in, PT := #v_pt, Q => #v_q, ET => #v_et);
END_FUNCTION_BLOCK

FUNCTION_BLOCK "FB_Scl_sl006"   // FB28, SCL
{ S7_Optimized_Access := 'TRUE' }
VERSION : 0.1
   VAR_INPUT
      v_in : Bool;
      v_r : Bool;
      v_pt : Time;
   END_VAR
   VAR_OUTPUT
      v_q : Bool;
      v_et : Time;
   END_VAR
   VAR
      inst : TONR_TIME;
   END_VAR
BEGIN
   #inst(IN := #v_in, R := #v_r, PT := #v_pt, Q => #v_q, ET => #v_et);
END_FUNCTION_BLOCK

FUNCTION_BLOCK "FB_Scl_sl015"   // FB29, SCL
{ S7_Optimized_Access := 'TRUE' }
VERSION : 0.1
   VAR_INPUT
      v_cd : Bool;
      v_ld : Bool;
      v_pv : Int;
   END_VAR
   VAR_OUTPUT
      v_q : Bool;
      v_cv : Char;
   END_VAR
   VAR
      inst : CTD_INT;
   END_VAR
BEGIN
   #inst(CD := #v_cd, LD := #v_ld, PV := #v_pv, Q => #v_q, CV => #v_cv);
END_FUNCTION_BLOCK

FUNCTION_BLOCK "FB_Scl_sl016"   // FB30, SCL
{ S7_Optimized_Access := 'TRUE' }
VERSION : 0.1
   VAR_INPUT
      v_cu : Bool;
      v_cd : Bool;
      v_r : Bool;
      v_ld : Bool;
      v_pv : Int;
   END_VAR
   VAR_OUTPUT
      v_qu : Bool;
      v_qd : Bool;
      v_cv : Char;
   END_VAR
   VAR
      inst : CTUD_INT;
   END_VAR
BEGIN
   #inst(CU := #v_cu, CD := #v_cd, R := #v_r, LD := #v_ld, PV := #v_pv, QU => #v_qu, QD => #v_qd, CV => #v_cv);
END_FUNCTION_BLOCK

FUNCTION_BLOCK "FB_Scl_sl053"   // FB31, SCL
{ S7_Optimized_Access := 'TRUE' }
VERSION : 0.1
   VAR_INPUT
      v_req : Bool;
      v_db : DB_ANY;
      v_index : DInt;
   END_VAR
   VAR_OUTPUT
      v_busy : Bool;
      v_done : Bool;
      v_error : Int;
   END_VAR
   VAR_IN_OUT
      v_value : Variant;
   END_VAR
   VAR
      inst : ReadFromArrayDBL;
   END_VAR
BEGIN
   #inst(req := #v_req, db := #v_db, index := #v_index, value := #v_value, busy => #v_busy, done => #v_done, error => #v_error);
END_FUNCTION_BLOCK

FUNCTION_BLOCK "FB_Scl_sl054"   // FB32, SCL
{ S7_Optimized_Access := 'TRUE' }
VERSION : 0.1
   VAR_INPUT
      v_req : Bool;
      v_db : DB_ANY;
      v_index : DInt;
      v_value : Variant;
   END_VAR
   VAR_OUTPUT
      v_busy : Bool;
      v_done : Bool;
      v_error : Int;
   END_VAR
   VAR
      inst : WriteToArrayDBL;
   END_VAR
BEGIN
   #inst(req := #v_req, db := #v_db, index := #v_index, value := #v_value, busy => #v_busy, done => #v_done, error => #v_error);
END_FUNCTION_BLOCK

FUNCTION_BLOCK "FB_Scl_sl058"   // FB33, SCL
{ S7_Optimized_Access := 'TRUE' }
VERSION : 0.1
   VAR_INPUT
      v_area : Byte;
      v_dbnumber : DInt;
      v_byteoffset : DInt;
      v_bitoffset : Int;
      v_value : Bool;
   END_VAR
BEGIN
   POKE_BOOL(area := #v_area, dbNumber := #v_dbnumber, byteOffset := #v_byteoffset, bitOffset := #v_bitoffset, value := #v_value);
END_FUNCTION_BLOCK

FUNCTION_BLOCK "FB_Scl_sl059"   // FB34, SCL
{ S7_Optimized_Access := 'TRUE' }
VERSION : 0.1
   VAR_INPUT
      v_area_src : Byte;
      v_dbnumber_src : DInt;
      v_byteoffset_src : DInt;
      v_area_dest : Byte;
      v_dbnumber_dest : DInt;
      v_byteoffset_dest : DInt;
      v_count : DInt;
   END_VAR
BEGIN
   POKE_BLK(area_src := #v_area_src, dbNumber_src := #v_dbnumber_src, byteOffset_src := #v_byteoffset_src, area_dest := #v_area_dest, dbNumber_dest := #v_dbnumber_dest, byteOffset_dest := #v_byteoffset_dest, count := #v_count);
END_FUNCTION_BLOCK

FUNCTION_BLOCK "FB_Scl_sl064"   // FB35, SCL
{ S7_Optimized_Access := 'TRUE' }
VERSION : 0.1
   VAR_INPUT
      v_src : Variant;
   END_VAR
   VAR_OUTPUT
      v_dst : Date;
   END_VAR
BEGIN
   VariantGet(SRC := #v_src, DST => #v_dst);
END_FUNCTION_BLOCK

FUNCTION_BLOCK "FB_Scl_sl065"   // FB36, SCL
{ S7_Optimized_Access := 'TRUE' }
VERSION : 0.1
   VAR_INPUT
      v_src : Date;
      v_dst : Variant;
   END_VAR
BEGIN
   VariantPut(SRC := #v_src, DST := #v_dst);
END_FUNCTION_BLOCK

FUNCTION_BLOCK "FB_Scl_sl009"   // FB37, SCL
{ S7_Optimized_Access := 'TRUE' }
VERSION : 0.1
   VAR_INPUT
      v_t_no : Timer;
      v_s : Bool;
      v_tv : S5Time;
      v_r : Bool;
   END_VAR
   VAR_OUTPUT
      v_q : Bool;
      v_bi : Word;
   END_VAR
BEGIN
   #v_bi := S_PULSE(T_NO := #v_t_no, S := #v_s, TV := #v_tv, R := #v_r, Q => #v_q);
END_FUNCTION_BLOCK

FUNCTION_BLOCK "FB_Scl_sl024"   // FB38, SCL
{ S7_Optimized_Access := 'TRUE' }
VERSION : 0.1
   VAR_INPUT
      v_in : SInt;
   END_VAR
   VAR_OUTPUT
      v_ret : SInt;
   END_VAR
BEGIN
   #v_ret := ABS(IN := #v_in);
END_FUNCTION_BLOCK

FUNCTION_BLOCK "FB_Scl_sl025"   // FB39, SCL
{ S7_Optimized_Access := 'TRUE' }
VERSION : 0.1
   VAR_INPUT
      v_in1 : Time;
      v_in2 : Time;
   END_VAR
   VAR_OUTPUT
      v_ret : Time;
   END_VAR
BEGIN
   #v_ret := MIN(IN1 := #v_in1, IN2 := #v_in2);
END_FUNCTION_BLOCK

FUNCTION_BLOCK "FB_Scl_sl026"   // FB40, SCL
{ S7_Optimized_Access := 'TRUE' }
VERSION : 0.1
   VAR_INPUT
      v_in1 : Time;
      v_in2 : Time;
   END_VAR
   VAR_OUTPUT
      v_ret : Time;
   END_VAR
BEGIN
   #v_ret := MAX(IN1 := #v_in1, IN2 := #v_in2);
END_FUNCTION_BLOCK

FUNCTION_BLOCK "FB_Scl_sl038"   // FB41, SCL
{ S7_Optimized_Access := 'TRUE' }
VERSION : 0.1
   VAR_INPUT
      v_in : Real;
   END_VAR
   VAR_OUTPUT
      v_ret : Real;
   END_VAR
BEGIN
   #v_ret := FRAC(IN := #v_in);
END_FUNCTION_BLOCK

FUNCTION_BLOCK "FB_Scl_sl010"   // FB42, SCL
{ S7_Optimized_Access := 'TRUE' }
VERSION : 0.1
   VAR_INPUT
      v_t_no : Timer;
      v_s : Bool;
      v_tv : S5Time;
      v_r : Bool;
   END_VAR
   VAR_OUTPUT
      v_q : Bool;
      v_bi : Word;
   END_VAR
BEGIN
   #v_bi := S_PEXT(T_NO := #v_t_no, S := #v_s, TV := #v_tv, R := #v_r, Q => #v_q);
END_FUNCTION_BLOCK

FUNCTION_BLOCK "FB_Scl_sl011"   // FB43, SCL
{ S7_Optimized_Access := 'TRUE' }
VERSION : 0.1
   VAR_INPUT
      v_t_no : Timer;
      v_s : Bool;
      v_tv : S5Time;
      v_r : Bool;
   END_VAR
   VAR_OUTPUT
      v_q : Bool;
      v_bi : Word;
   END_VAR
BEGIN
   #v_bi := S_ODT(T_NO := #v_t_no, S := #v_s, TV := #v_tv, R := #v_r, Q => #v_q);
END_FUNCTION_BLOCK

FUNCTION_BLOCK "FB_Scl_sl012"   // FB44, SCL
{ S7_Optimized_Access := 'TRUE' }
VERSION : 0.1
   VAR_INPUT
      v_t_no : Timer;
      v_s : Bool;
      v_tv : S5Time;
      v_r : Bool;
   END_VAR
   VAR_OUTPUT
      v_q : Bool;
      v_bi : Word;
   END_VAR
BEGIN
   #v_bi := S_ODTS(T_NO := #v_t_no, S := #v_s, TV := #v_tv, R := #v_r, Q => #v_q);
END_FUNCTION_BLOCK

FUNCTION_BLOCK "FB_Scl_sl013"   // FB45, SCL
{ S7_Optimized_Access := 'TRUE' }
VERSION : 0.1
   VAR_INPUT
      v_t_no : Timer;
      v_s : Bool;
      v_tv : S5Time;
      v_r : Bool;
   END_VAR
   VAR_OUTPUT
      v_q : Bool;
      v_bi : Word;
   END_VAR
BEGIN
   #v_bi := S_OFFDT(T_NO := #v_t_no, S := #v_s, TV := #v_tv, R := #v_r, Q => #v_q);
END_FUNCTION_BLOCK

FUNCTION_BLOCK "FB_Scl_sl017"   // FB46, SCL
{ S7_Optimized_Access := 'TRUE' }
VERSION : 0.1
   VAR_INPUT
      v_c_no : Counter;
      v_cu : Bool;
      v_s : Bool;
      v_pv : Word;
      v_r : Bool;
   END_VAR
   VAR_OUTPUT
      v_q : Bool;
      v_cv : Word;
   END_VAR
BEGIN
   #v_cv := S_CU(C_NO := #v_c_no, CU := #v_cu, S := #v_s, PV := #v_pv, R := #v_r, Q => #v_q);
END_FUNCTION_BLOCK

FUNCTION_BLOCK "FB_Scl_sl018"   // FB47, SCL
{ S7_Optimized_Access := 'TRUE' }
VERSION : 0.1
   VAR_INPUT
      v_c_no : Counter;
      v_cd : Bool;
      v_s : Bool;
      v_pv : Word;
      v_r : Bool;
   END_VAR
   VAR_OUTPUT
      v_q : Bool;
      v_cv : Word;
   END_VAR
BEGIN
   #v_cv := S_CD(C_NO := #v_c_no, CD := #v_cd, S := #v_s, PV := #v_pv, R := #v_r, Q => #v_q);
END_FUNCTION_BLOCK

FUNCTION_BLOCK "FB_Scl_sl019"   // FB48, SCL
{ S7_Optimized_Access := 'TRUE' }
VERSION : 0.1
   VAR_INPUT
      v_c_no : Counter;
      v_cu : Bool;
      v_cd : Bool;
      v_s : Bool;
      v_pv : Word;
      v_r : Bool;
   END_VAR
   VAR_OUTPUT
      v_q : Bool;
      v_cv : Word;
   END_VAR
BEGIN
   #v_cv := S_CUD(C_NO := #v_c_no, CU := #v_cu, CD := #v_cd, S := #v_s, PV := #v_pv, R := #v_r, Q => #v_q);
END_FUNCTION_BLOCK

FUNCTION_BLOCK "FB_Scl_sl027"   // FB49, SCL
{ S7_Optimized_Access := 'TRUE' }
VERSION : 0.1
   VAR_INPUT
      v_mn : Time;
      v_in : Time;
      v_mx : Time;
   END_VAR
   VAR_OUTPUT
      v_ret : Time;
   END_VAR
BEGIN
   #v_ret := LIMIT(MN := #v_mn, IN := #v_in, MX := #v_mx);
END_FUNCTION_BLOCK

FUNCTION_BLOCK "FB_Scl_sl028"   // FB50, SCL
{ S7_Optimized_Access := 'TRUE' }
VERSION : 0.1
   VAR_INPUT
      v_in : Real;
   END_VAR
   VAR_OUTPUT
      v_ret : Real;
   END_VAR
BEGIN
   #v_ret := SQR(IN := #v_in);
END_FUNCTION_BLOCK

FUNCTION_BLOCK "FB_Scl_sl029"   // FB51, SCL
{ S7_Optimized_Access := 'TRUE' }
VERSION : 0.1
   VAR_INPUT
      v_in : Real;
   END_VAR
   VAR_OUTPUT
      v_ret : Real;
   END_VAR
BEGIN
   #v_ret := SQRT(IN := #v_in);
END_FUNCTION_BLOCK

FUNCTION_BLOCK "FB_Scl_sl030"   // FB52, SCL
{ S7_Optimized_Access := 'TRUE' }
VERSION : 0.1
   VAR_INPUT
      v_in : Real;
   END_VAR
   VAR_OUTPUT
      v_ret : Real;
   END_VAR
BEGIN
   #v_ret := LN(IN := #v_in);
END_FUNCTION_BLOCK

FUNCTION_BLOCK "FB_Scl_sl031"   // FB53, SCL
{ S7_Optimized_Access := 'TRUE' }
VERSION : 0.1
   VAR_INPUT
      v_in : Real;
   END_VAR
   VAR_OUTPUT
      v_ret : Real;
   END_VAR
BEGIN
   #v_ret := EXP(IN := #v_in);
END_FUNCTION_BLOCK

FUNCTION_BLOCK "FB_Scl_sl032"   // FB54, SCL
{ S7_Optimized_Access := 'TRUE' }
VERSION : 0.1
   VAR_INPUT
      v_in : Real;
   END_VAR
   VAR_OUTPUT
      v_ret : Real;
   END_VAR
BEGIN
   #v_ret := SIN(IN := #v_in);
END_FUNCTION_BLOCK

FUNCTION_BLOCK "FB_Scl_sl033"   // FB55, SCL
{ S7_Optimized_Access := 'TRUE' }
VERSION : 0.1
   VAR_INPUT
      v_in : Real;
   END_VAR
   VAR_OUTPUT
      v_ret : Real;
   END_VAR
BEGIN
   #v_ret := COS(IN := #v_in);
END_FUNCTION_BLOCK

FUNCTION_BLOCK "FB_Scl_sl034"   // FB56, SCL
{ S7_Optimized_Access := 'TRUE' }
VERSION : 0.1
   VAR_INPUT
      v_in : Real;
   END_VAR
   VAR_OUTPUT
      v_ret : Real;
   END_VAR
BEGIN
   #v_ret := TAN(IN := #v_in);
END_FUNCTION_BLOCK

FUNCTION_BLOCK "FB_Scl_sl035"   // FB57, SCL
{ S7_Optimized_Access := 'TRUE' }
VERSION : 0.1
   VAR_INPUT
      v_in : Real;
   END_VAR
   VAR_OUTPUT
      v_ret : Real;
   END_VAR
BEGIN
   #v_ret := ASIN(IN := #v_in);
END_FUNCTION_BLOCK

FUNCTION_BLOCK "FB_Scl_sl036"   // FB58, SCL
{ S7_Optimized_Access := 'TRUE' }
VERSION : 0.1
   VAR_INPUT
      v_in : Real;
   END_VAR
   VAR_OUTPUT
      v_ret : Real;
   END_VAR
BEGIN
   #v_ret := ACOS(IN := #v_in);
END_FUNCTION_BLOCK

FUNCTION_BLOCK "FB_Scl_sl037"   // FB59, SCL
{ S7_Optimized_Access := 'TRUE' }
VERSION : 0.1
   VAR_INPUT
      v_in : Real;
   END_VAR
   VAR_OUTPUT
      v_ret : Real;
   END_VAR
BEGIN
   #v_ret := ATAN(IN := #v_in);
END_FUNCTION_BLOCK

FUNCTION_BLOCK "FB_Scl_sl039"   // FB60, SCL
{ S7_Optimized_Access := 'TRUE' }
VERSION : 0.1
   VAR_INPUT
      v_src_array : Byte;
   END_VAR
   VAR_OUTPUT
      v_ret : Byte;
   END_VAR
   VAR_IN_OUT
      v_dest_variable : Variant;
      v_pos : DInt;
   END_VAR
BEGIN
   #v_ret := Deserialize(SRC_ARRAY := #v_src_array, DEST_VARIABLE => #v_dest_variable, POS := #v_pos);
END_FUNCTION_BLOCK

FUNCTION_BLOCK "FB_Scl_sl050"   // FB61, SCL
{ S7_Optimized_Access := 'TRUE' }
VERSION : 0.1
   VAR_INPUT
      v_in : Word;
   END_VAR
   VAR_OUTPUT
      v_ret : Word;
   END_VAR
BEGIN
   #v_ret := SWAP(IN := #v_in);
END_FUNCTION_BLOCK

FUNCTION_BLOCK "FB_Scl_sl055"   // FB62, SCL
{ S7_Optimized_Access := 'TRUE' }
VERSION : 0.1
   VAR_INPUT
      v_area : Byte;
      v_dbnumber : DInt;
      v_byteoffset : DInt;
   END_VAR
   VAR_OUTPUT
      v_ret : Byte;
   END_VAR
BEGIN
   #v_ret := PEEK(area := #v_area, dbNumber := #v_dbnumber, byteOffset := #v_byteoffset);
END_FUNCTION_BLOCK

FUNCTION_BLOCK "FB_Scl_sl073"   // FB63, SCL
{ S7_Optimized_Access := 'TRUE' }
VERSION : 0.1
   VAR_INPUT
      v_in : Real;
   END_VAR
   VAR_OUTPUT
      v_ret : Real;
   END_VAR
BEGIN
   #v_ret := ROUND(IN := #v_in);
END_FUNCTION_BLOCK

FUNCTION_BLOCK "FB_Scl_sl074"   // FB64, SCL
{ S7_Optimized_Access := 'TRUE' }
VERSION : 0.1
   VAR_INPUT
      v_in : Real;
   END_VAR
   VAR_OUTPUT
      v_ret : Real;
   END_VAR
BEGIN
   #v_ret := CEIL(IN := #v_in);
END_FUNCTION_BLOCK

FUNCTION_BLOCK "FB_Scl_sl075"   // FB65, SCL
{ S7_Optimized_Access := 'TRUE' }
VERSION : 0.1
   VAR_INPUT
      v_in : Real;
   END_VAR
   VAR_OUTPUT
      v_ret : Real;
   END_VAR
BEGIN
   #v_ret := FLOOR(IN := #v_in);
END_FUNCTION_BLOCK

FUNCTION_BLOCK "FB_Scl_sl076"   // FB66, SCL
{ S7_Optimized_Access := 'TRUE' }
VERSION : 0.1
   VAR_INPUT
      v_in : Real;
   END_VAR
   VAR_OUTPUT
      v_ret : Real;
   END_VAR
BEGIN
   #v_ret := TRUNC(IN := #v_in);
END_FUNCTION_BLOCK

FUNCTION_BLOCK "FB_Scl_sl077"   // FB67, SCL
{ S7_Optimized_Access := 'TRUE' }
VERSION : 0.1
   VAR_INPUT
      v_min : Real;
      v_value : Real;
      v_max : Real;
   END_VAR
   VAR_OUTPUT
      v_ret : Real;
   END_VAR
BEGIN
   #v_ret := SCALE_X(MIN := #v_min, VALUE := #v_value, MAX := #v_max);
END_FUNCTION_BLOCK

FUNCTION_BLOCK "FB_Scl_sl078"   // FB68, SCL
{ S7_Optimized_Access := 'TRUE' }
VERSION : 0.1
   VAR_INPUT
      v_min : Real;
      v_value : Real;
      v_max : Real;
   END_VAR
   VAR_OUTPUT
      v_ret : Real;
   END_VAR
BEGIN
   #v_ret := NORM_X(MIN := #v_min, VALUE := #v_value, MAX := #v_max);
END_FUNCTION_BLOCK

FUNCTION_BLOCK "FB_Fbd_ex005"   // FB69, FBD
{ S7_Optimized_Access := 'TRUE' }
   VAR_INPUT
      v_in1 : DTL;
      v_in2 : DTL;
   END_VAR
   VAR_OUTPUT
      v_out : Time;
   END_VAR
BEGIN

REGION Network 1: T_DIFF - Time difference
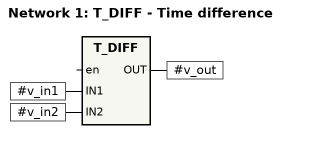
   #v_out := T_DIFF(IN1 := #v_in1, IN2 := #v_in2);
END_REGION
END_FUNCTION_BLOCK

FUNCTION_BLOCK "FB_Fbd_ex007"   // FB70, FBD
{ S7_Optimized_Access := 'TRUE' }
   VAR_INPUT
      v_in : DTL;
   END_VAR
   VAR_OUTPUT
      v_ret_val : Int;
   END_VAR
BEGIN

REGION Network 1: WR_SYS_T - Set time-of-day
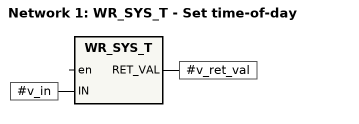
   #v_ret_val := WR_SYS_T(IN := #v_in);
END_REGION
END_FUNCTION_BLOCK

FUNCTION_BLOCK "FB_Fbd_ex008"   // FB71, FBD
{ S7_Optimized_Access := 'TRUE' }
   VAR_OUTPUT
      v_ret_val : Int;
      v_out : DTL;
   END_VAR
BEGIN

REGION Network 1: RD_SYS_T - Read time-of-day
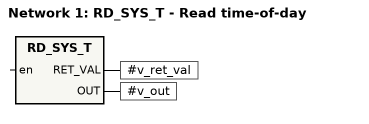
   #v_ret_val := RD_SYS_T(OUT => #v_out);
END_REGION
END_FUNCTION_BLOCK

FUNCTION_BLOCK "FB_Fbd_ex009"   // FB72, FBD
{ S7_Optimized_Access := 'TRUE' }
   VAR_OUTPUT
      v_ret_val : Int;
      v_out : DTL;
   END_VAR
BEGIN

REGION Network 1: RD_LOC_T - Read local time
